// TIA Portal V20 export
TYPE "WT3_Verdampfer_Status_UDT"
   STRUCT
      iHandshake : Int;
      Alarm : Struct
         bE0000_KonfigAlarm : Bool;
         bE0001_Reserviert : Bool;
         bE0002_InvUngueltig : Bool;
         bE0003_Reserviert : Bool;
         bE0004_FrostschutzFehler : Bool;
         bE0005_VerdampferpumpeAlarmBetrieb : Bool;
         bE0006_VerdampferpumpeAlarmStillstand : Bool;
         bE0007_VerdampferEintrittWarm : Bool;
         bE0008_NiveauAbscheiderHochFehler : Bool;
         bE0009_KonfigAlarmUmstellungDIPolarität : Bool;
         bE0010_Reserviert : Bool;
         bE0011_Reserviert : Bool;
         bE0012_NiveauAbscheider2HochAlarm : Bool;
         bE0013_KonfigAlarmÖlrektifizierung : Bool;
         bE0014_Reserviert : Bool;
         bE0015_Reserviert : Bool;
         bE0016_MediumüberdruckZuTief : Bool;
         bE0017_KonfigAlarmEERVerdichter : Bool;
         bE0018_DurchflussstörungVerdampferInBetrieb : Bool;
         bE0019_DurchflussstörungVerdampferBeimStart : Bool;
         bE0020_DurchflussstörungVerdampferImStillstand : Bool;
         bE0021_Reserviert : Bool;
         bE0022_Strömungsaufbau : Bool;
         bE0023_StrömungImBetrieb : Bool;
         bE0024_StrömungImStillstand : Bool;
         b051_Reserve : Bool;
         b052_Reserve : Bool;
         b053_Reserve : Bool;
         b054_Reserve : Bool;
         b055_Reserve : Bool;
         bE0030_AbsperrklappeEintrittNichtOffen : Bool;
         bE0031_AbsperrklappeEintrittNichtZu : Bool;
         bE0032_AbsperrklappeAustrittNichtOffen : Bool;
         bE0033_AbsperrklappeAustrittNichtZu : Bool;
         bE0034_NH3inSekundärkreis : Bool;
         bE0035_StörungRegelventilAbscheider1 : Bool;
         bE0036_StörungRegelventilAbscheider2 : Bool;
         bE0337_ExternFehler : Bool;
         b066_Reserve : Bool;
         b067_Reserve : Bool;
         by07_Reserve : Byte;
         by08_Reserve : Byte;
         by09_Reserve : Byte;
         by10_Reserve : Byte;
         by11_Reserve : Byte;
         by12_Reserve : Byte;
         by13_Reserve : Byte;
         by14_Reserve : Byte;
         by15_Reserve : Byte;
         by16_Reserve : Byte;
         by17_Reserve : Byte;
         by18_Reserve : Byte;
         by19_Reserve : Byte;
         by20_Reserve : Byte;
         by21_Reserve : Byte;
         by22_Reserve : Byte;
         by23_Reserve : Byte;
         by24_Reserve : Byte;
         by25_Reserve : Byte;
         by26_Reserve : Byte;
         bE0200_AlarmKabelbruch : Bool;
         b271_Reserve : Bool;
         b272_Reserve : Bool;
         b273_Reserve : Bool;
         b274_Reserve : Bool;
         b275_Reserve : Bool;
         b276_Reserve : Bool;
         b277_Reserve : Bool;
         by28_Reserve : Byte;
         by29_Reserve : Byte;
         by30_Reserve : Byte;
         by31_Reserve : Byte;
         by32_Reserve : Byte;
         by33_Reserve : Byte;
      END_STRUCT;
      Warnung : Struct
         bA1000_Reserviert : Bool;
         bA1001_SlaveAusg : Bool;
         bA1002_Reserviert : Bool;
         bA1003_HauptMasterAusg : Bool;
         bA1004_Reserviert : Bool;
         bA1005_Reserviert : Bool;
         bA1006_Reserviert : Bool;
         bA1007_Reserviert : Bool;
         bA1008_Reserviert : Bool;
         bA1009_Reserviert : Bool;
         bA1010_MehrereVerdampferMasterAktiv : Bool;
         bA1011_ObjektIDMehrfVorhanden : Bool;
         bA1012_Reserviert : Bool;
         bA1013_Reserviert : Bool;
         bA1014_WarnungNiveauAbscheiderEndschalter : Bool;
         bA1015_WarnungNiveauAbscheider2Endschalter : Bool;
         bA1016_Reserviert : Bool;
         bA1017_Reserviert : Bool;
         bA1018_Reserviert : Bool;
         bA1019_Reserviert : Bool;
         bA1020_Reserviert : Bool;
         bA1021_ÖlSensorFunktionsstörung : Bool;
         bA1022_Reserviert : Bool;
         bA1023_Reserviert : Bool;
         bA1024_Reserviert : Bool;
         bA1025_ÖlrektifizierungLaufzeit : Bool;
         bA1026_TÖlsammlerSollNichtErreicht : Bool;
         bA1027_ÖlSammlerNiveauZuTief : Bool;
         bA1028_TÖlSammlerZuHoch : Bool;
         bA1029_TÖlSammlerZuTief : Bool;
         b376_Reserve : Bool;
         b377_Reserve : Bool;
         by38_Reserve : Byte;
         by39_Reserve : Byte;
         by40_Reserve : Byte;
         by41_Reserve : Byte;
         by42_Reserve : Byte;
         by43_Reserve : Byte;
         by44_Reserve : Byte;
         by45_Reserve : Byte;
         by46_Reserve : Byte;
         by47_Reserve : Byte;
         by48_Reserve : Byte;
         by49_Reserve : Byte;
         by50_Reserve : Byte;
         by51_Reserve : Byte;
         by52_Reserve : Byte;
         by53_Reserve : Byte;
         by54_Reserve : Byte;
         by55_Reserve : Byte;
         by56_Reserve : Byte;
         by57_Reserve : Byte;
         by58_Reserve : Byte;
         bA1200_WarnungKabelbruch : Bool;
         b591_Reserve : Bool;
         b592_Reserve : Bool;
         b593_Reserve : Bool;
         b594_Reserve : Bool;
         b595_Reserve : Bool;
         b596_Reserve : Bool;
         b597_Reserve : Bool;
         by60_Reserve : Byte;
         by61_Reserve : Byte;
         by62_Reserve : Byte;
         by63_Reserve : Byte;
         by64_Reserve : Byte;
         by65_Reserve : Byte;
      END_STRUCT;
      Zustand : Struct
         bAlarmzustandAktiv : Bool;
         bWarnzustandAktiv : Bool;
         bSystemMeldungAktiv : Bool;
         bSeviceMeldungAktiv : Bool;
         bStopManuell : Bool;
         bStopAuto : Bool;
         bStopExtern : Bool;
         bBetriebAuto : Bool;
         bBetriebManuell : Bool;
         bAnlaufAuto : Bool;
         bAnlaufManuell : Bool;
         bManuellStoppen : Bool;
         b674_Reserve : Bool;
         b675_Reserve : Bool;
         b676_Reserve : Bool;
         b677_Reserve : Bool;
         by68_Reserve : Byte;
         by69_Reserve : Byte;
         bInventarAufnahme : Bool;
         b701_Reserve : Bool;
         bStandbyMasterInit : Bool;
         bStandbyMasterPassiv : Bool;
         bStandbyMasterAktiv : Bool;
         bMasterGesperrt : Bool;
         bSollwertAbsenkung : Bool;
         bIstwertVentilfühler : Bool;
         bIstwertPSaug : Bool;
         bVerdampferpumpeManuell : Bool;
         bAbsperrklappenOeffnen : Bool;
         bAbsperrklappenSchliessen : Bool;
         bSpülungAktiv : Bool;
         b715_Reserve : Bool;
         b716_Reserve : Bool;
         b717_Reserve : Bool;
         by72_Reserve : Byte;
         by73_Reserve : Byte;
         by74_Reserve : Byte;
         by75_Reserve : Byte;
         by76_Reserve : Byte;
         by77_Reserve : Byte;
         by78_Reserve : Byte;
         by79_Reserve : Byte;
         by80_Reserve : Byte;
         by81_Reserve : Byte;
      END_STRUCT;
      "Allgemeine Meldungen" : Struct
         b4000_AllgemeineMeldung_1 : Bool;
         b4001_AllgemeineMeldung_2 : Bool;
         b4002_AllgemeineMeldung_3 : Bool;
         b4003_AllgemeineMeldung_4 : Bool;
         b4004_AllgemeineMeldung_5 : Bool;
         b4005_AllgemeineMeldung_6 : Bool;
         b4006_AllgemeineMeldung_7 : Bool;
         b4007_AllgemeineMeldung_8 : Bool;
         by83_Reserve : Byte;
         by84_Reserve : Byte;
         by85_Reserve : Byte;
      END_STRUCT;
      DigIn : Struct
         bSollwertB : Bool;
         bRückmeldungVerdampferpumpe : Bool;
         btKühlstelleDigital : Bool;
         bStartbefehlKühlstelle : Bool;
         bAbscheiderNiveauHoch : Bool;
         bAbscheiderNiveauregFreigabe : Bool;
         bAbscheider2NiveauHoch : Bool;
         bAbscheider2NiveauregFreigabe : Bool;
         bAbscheiderBetriebsart : Bool;
         bAbscheider2Betriebsart : Bool;
         bAbscheiderNiveauEndschalterOffen : Bool;
         bAbscheiderNiveauEndschalterGeschlossen : Bool;
         bAbscheider2NiveauEndschalterOffen : Bool;
         bAbscheider2NiveauEndschalterGeschlossen : Bool;
         bFrostschutzDigital : Bool;
         bMediumKreislÜberdruck : Bool;
         bÖlSensorÖlrektifizierung : Bool;
         bStrömungswächter : Bool;
         bNiveauTiefÖlsammler : Bool;
         bEndschalterAbsperrklappeEintrittOffen : Bool;
         bEndschalterAbsperrklappeEintrittZu : Bool;
         bEndschalterAbsperrklappeAustrittOffen : Bool;
         bEndschalterAbsperrklappeAustrittZu : Bool;
         bNH3AlarmSekunkdärkreis : Bool;
         by89_Reserve : Byte;
         by90_Reserve : Byte;
         by91_Reserve : Byte;
         by92_Reserve : Byte;
         by93_Reserve : Byte;
      END_STRUCT;
      DigOut : Struct
         bStratbefehlVerdampferpumpe : Bool;
         bMVKühlstelle : Bool;
         bAbscheiderNiveauregelung : Bool;
         bAbscheider2Niveauregelung : Bool;
         bMVAbscheiderNachspeisung : Bool;
         bMVAbscheider2Nachspeisung : Bool;
         bÖlrektifizierung : Bool;
         bÖlzulauf : Bool;
         bÖlsammlerHeizung : Bool;
         bDruckbeaufschlagung : Bool;
         bDruckbeaufschlagungHD : Bool;
         bDruckbeaufschlagungND : Bool;
         bMvEntgasungOelsammler : Bool;
         bMvEntgasungOelsammelrohr : Bool;
         bAbsperrklappeEintritt : Bool;
         bAbsperrklappeAustritt : Bool;
         by96_Reserve : Byte;
         by97_Reserve : Byte;
         by98_Reserve : Byte;
         by99_Reserve : Byte;
         by100_Reserve : Byte;
         by101_Reserve : Byte;
      END_STRUCT;
      ch1021_Reserve : Char;
      chVerdReglerEinheit : Char;
      rVerdReglerIstwert : Real;
      rVerdReglerSollwert : Real;
      rVerdReglerAusgang : Real;
      rVerdEintrittstemperatur : Real;
      rVerdAustrittstemperatur : Real;
      diStatusSollwertrampe : DInt;
      rVerdReglerAusgang2 : Real;
      rVerdPumpe : Real;
      rVerddreiwegventil : Real;
      rTVentlfühler : Real;
      rFrostschutzFühler : Real;
      rTKühlstelle : Real;
      rAbscheiderNiveau : Real;
      rAbscheiderNiveauregelung : Real;
      rAbscheiderNiveau2 : Real;
      rAbscheiderNiveauregelung2 : Real;
      rPSaugseiteBar : Real;
      rPSaugseiteTemp : Real;
      rÜberströmventil : Real;
      rVolumenstrom : Real;
      rThermischeLeistung : Real;
      rEERVerdichter : Real;
      rEERAnlage : Real;
      rMediumKreislÜberdruck : Real;
      rAuxAnalog1 : Real;
      rAuxAnalog2 : Real;
      rTÖlsammler : Real;
      rTGradientBegrenzung : Real;
      rAuxAnalog3 : Real;
      rAuxAnalog4 : Real;
      byReserve : Array[224..629] of Byte;
   END_STRUCT;
END_TYPE
